(* IEC 61131-3 sources: PLCCodeForge/Autothink.UIA/Docs/Samples, 1 file *)

(* ---- program_demo.st ---- *)
PROGRAM Main
VAR
    counter : INT := 0;
END_VAR

counter := counter + 1;
END_PROGRAM
